(* IEC 61131-3 sources: rusty/compiler/plc_cfc/fixtures/blocks/invalid/function_duplicate_return, 1 file *)

(* ---- myAdd.st ---- *)
FUNCTION myAdd : DINT
VAR_INPUT
    in1 : DINT;
    in2 : DINT;
END_VAR
    myAdd := in1 + in2;
END_FUNCTION
